(* IEC 61131-3 sources: Test-Git_ESME26/TestProgettoESME_26.fbsproj/PacDriveLib_Motion_Migration_Example.device.xml.v3^/Plc Logic.plclogic.xml.v3^/Application.application.xml.v3^/Sercos_PacDriveLib/WriteIDN, 2 files *)

(* ---- FC_SercosWriteIDN.fn.st ---- *)
FUNCTION FC_SercosWriteIDN : DINT
VAR_INPUT
	i_uiTopoAddr : UINT;
	i_etSercosParameterType : ET_SercosParameterType;
	i_uiIDN : UINT;
	i_etWriteIDNType : ET_SercosWriteIDNType;
	i_dwValue : DWORD;
END_VAR
VAR
	dwIDN : DWORD;
	dwValue : DWORD;
END_VAR

dwValue := i_dwValue;

IF i_etSercosParameterType = ET_SercosParameterType.S_Parameter THEN
	dwIDN := i_uiIDN;
ELSE
	dwIDN := 16#8000 + i_uiIDN;
END_IF

FC_SercosWriteIDN := SMM6xx.FC_SercosWriteServiceDataByTopAddr(
	i_wTopoAddr := i_uiTopoAddr,
	i_dwIDN := dwIDN,
	i_wType := TO_UINT(i_etWriteIDNType),
	i_lwPointerToData := TO_LWORD(ADR(dwValue)),
	i_wMaxDataLen := 2);

(* ---- FB_Set230VModeAsync.fb.st ---- *)
FUNCTION_BLOCK FB_Set230VModeAsync IMPLEMENTS SE_Async.IF_Async
VAR_INPUT
	i_ifSercosIdentificationAccess : SDI.IF_SercosIdentificationAccess;
END_VAR
VAR_OUTPUT
	q_diResult : DINT;
	q_sDiagMsg : STRING[255];
END_VAR
VAR
	xDone_loc : Bool;
END_VAR
